// TIA Portal V21 export
// export: Created 2026-11-07T15:24:55.5957561Z, ExportSetting WithDefaults, DisplayName Totally Integrated Automation Portal, DisplayVersion V21, DisplayName STEP 7 Professional, DisplayVersion V21, DisplayName STEP 7 Safety, DisplayVersion V21, DisplayName Tech WebApplication, DisplayVersion V21, DisplayName WinCC Basic/Comfort/Advanced, DisplayVersion V21, DisplayName WinCC Unified, DisplayVersion V21
Screen "R02_RectApp"  1024x768, Number=41, Template=Tpl
  ScreenLayer 
    Rectangle "P_CellRect" at 10,10 size 100x30  StyleItem=Rectangle
      RangeAppearanceAnimation "RangeAppearanceAnimation"
        tag P_Cell
        0..0: back #dedede, fore #000000
        1..1: back #a5a5a5, fore #000000
        2..2: back #8cafd7, fore #000000
        3..3: back #b9a0d2, fore #000000
        4..4: back #a5c8a5, fore #000000
        5..5: back #468ce6, fore #000000
        6..6: back #cdebff, fore #000000
        7..7: back #ffd700, fore #000000
